// Model of the TwinSAFE FB OR. Connected inputs are active.
// The Safety Editor refuses an OR with fewer than two OrIn ports connected: the model then reports
// Error with diagnostic bit 15 instead of running (see T_SafeFunctionBlockBase).
{attribute 'reflection'}
FUNCTION_BLOCK T_SafeOr EXTENDS T_SafeFunctionBlockBase
VAR_INPUT
    OrIn1 : BOOL;
    OrIn2 : BOOL;
    OrIn3 : BOOL;
    OrIn4 : BOOL;
    OrIn5 : BOOL;
    OrIn6 : BOOL;
    OrIn7 : BOOL;
    OrIn8 : BOOL;
    Parameters : ST_SafeLogicParameters;
END_VAR
VAR_OUTPUT
    OrOut : BOOL;
END_VAR
VAR
    {attribute 'is_connected' := 'OrIn1'}
    _orIn1Connected : BOOL;
    {attribute 'is_connected' := 'OrIn2'}
    _orIn2Connected : BOOL;
    {attribute 'is_connected' := 'OrIn3'}
    _orIn3Connected : BOOL;
    {attribute 'is_connected' := 'OrIn4'}
    _orIn4Connected : BOOL;
    {attribute 'is_connected' := 'OrIn5'}
    _orIn5Connected : BOOL;
    {attribute 'is_connected' := 'OrIn6'}
    _orIn6Connected : BOOL;
    {attribute 'is_connected' := 'OrIn7'}
    _orIn7Connected : BOOL;
    {attribute 'is_connected' := 'OrIn8'}
    _orIn8Connected : BOOL;
    _state : E_SafeFbState := E_SafeFbState.Stop;
END_VAR

SUPER^();

// At least two OrIn ports must be connected (Safety Editor: "OR does not have at least 2 input ports active and connected").
METHOD PROTECTED ConfigurationOk : BOOL
VAR
    connectedInputs : USINT;
END_VAR
connectedInputs := BOOL_TO_USINT(_orIn1Connected)
    + BOOL_TO_USINT(_orIn2Connected)
    + BOOL_TO_USINT(_orIn3Connected)
    + BOOL_TO_USINT(_orIn4Connected)
    + BOOL_TO_USINT(_orIn5Connected)
    + BOOL_TO_USINT(_orIn6Connected)
    + BOOL_TO_USINT(_orIn7Connected)
    + BOOL_TO_USINT(_orIn8Connected);

IF connectedInputs < 2 THEN
    _configurationFault := 'T_SafeOr: OR does not have at least 2 input ports active and connected';
    RETURN;
END_IF

ConfigurationOk := TRUE;
END_METHOD

METHOD PROTECTED Process
VAR
    result : BOOL;
END_VAR
result := FALSE;
result := result OR F_SafeInputValue(_orIn1Connected, Parameters.In1MakeContact, OrIn1);
result := result OR F_SafeInputValue(_orIn2Connected, Parameters.In2MakeContact, OrIn2);
result := result OR F_SafeInputValue(_orIn3Connected, Parameters.In3MakeContact, OrIn3);
result := result OR F_SafeInputValue(_orIn4Connected, Parameters.In4MakeContact, OrIn4);
result := result OR F_SafeInputValue(_orIn5Connected, Parameters.In5MakeContact, OrIn5);
result := result OR F_SafeInputValue(_orIn6Connected, Parameters.In6MakeContact, OrIn6);
result := result OR F_SafeInputValue(_orIn7Connected, Parameters.In7MakeContact, OrIn7);
result := result OR F_SafeInputValue(_orIn8Connected, Parameters.In8MakeContact, OrIn8);

IF NOT _fbRun THEN
    _state := E_SafeFbState.Stop;
ELSIF result THEN
    _state := E_SafeFbState.Run;
ELSE
    _state := E_SafeFbState.Safe;
END_IF

OrOut := (_state = E_SafeFbState.Run);
Error := FALSE;
Diag  := 0;
State := TO_BYTE(_state);
END_METHOD

END_FUNCTION_BLOCK

(* stored: Version 1.1.0.1
   POU T_SafeOr: Id {172c71ab-ec3d-5ccc-91c3-374336b4d74f}, SpecialFunc None
   Method ConfigurationOk: Id {b1fe103e-5756-4f48-95e1-ae3f8a72473d}
   Method Process: Id {6d72b5e1-d040-529f-8c8f-d3c7e840ffaf} *)
